PROGRAM main
  VAR
    rTemp : REAL;
    xAlarm : BOOL;
    xStart : BOOL;
  END_VAR

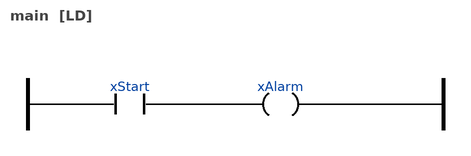
(* LD diagram, written out as Structured Text *)
xAlarm := xStart;
END_PROGRAM
